Yaskawa INFORM job: M_LONGP.JBI

/JOB
//NAME M_LONGP
//POS
///NPOS 0,0,0,0,0,0
//INST
<volatile>
///COMM Generated using RoboDK
///ATTR SC,RW
///GROUP1 RB1
NOP
CALL JOB:LONGPRO
CALL JOB:LONGPRO2
CALL JOB:LONGPRO3
CALL JOB:LONGPRO4
CALL JOB:LONGPRO5
END
